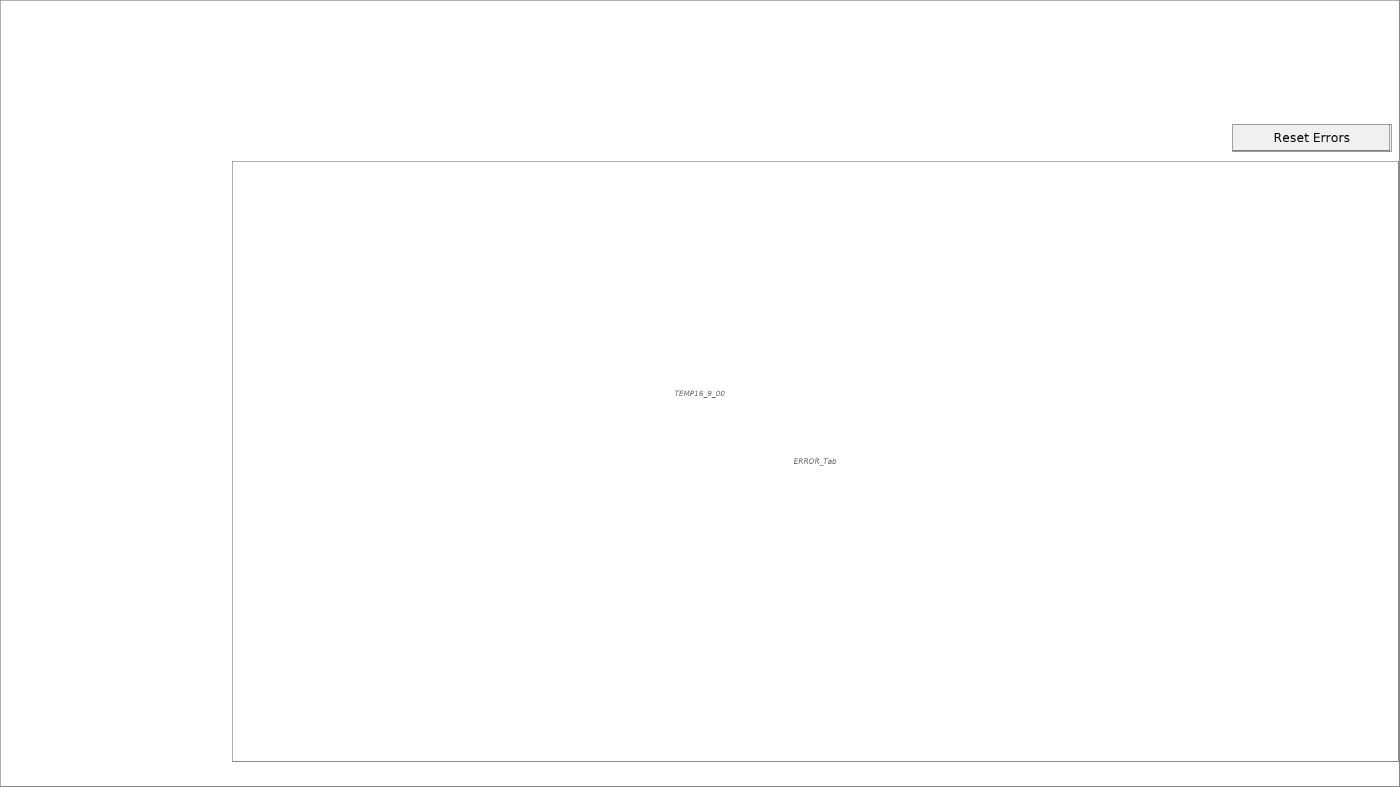
VISUALIZATION ERRORS_OPER_16_9  // 1920x1080
    Frame (0,0 1920x1080)
        shows TEMP16_9_00()
    Frame (318,221 1600x824)
        shows ERROR_Tab()
    Button (1690,170 218x38), "Reset Errors", pressed state: prg_Messages.ResetErrors
        toggle prg_Messages.ResetErrors
END_VISUALIZATION

(* stored: Version 1.1.0.1, ProductVersion 3.1.4024.13
   Visu ERRORS_OPER_16_9: Id {f1316b37-5571-4aeb-9cac-d7116779d41f} *)
